(* IEC 61131-3 sources: Versio-VersionControlSystem/fixtures/projects/TC3_PlcSample_reStrText/TC3_PlcSample_reStrText/LibraryDocumentationSample Project/LibPOUs/B_DocuElements/Images, 1 file *)

(* ---- FB_Libdoc_Images.st ---- *)
(*

**Absolute or relative file path as directive argument**

Absolute path

.. image:: C:\Tc3LibDocImages\tulpis.jpg
   :width: 70px

Relative path

.. image:: ../../LibPics/penguins.jpg
   :width: 70px

**Left aligned image**

.. image:: ../../LibPics/desert.jpg
   :width: 20%

Description of the function block. Description of the function block. Description of the function block.
Description of the function block. Description of the function block. Description of the function block.
Description of the function block. Description of the function block. Description of the function block.
Description of the function block. Description of the function block. Description of the function block.

**Floating image, left aligned**

.. image:: ../../LibPics/desert.jpg
   :width: 20%
   :align: left

Description of the function block. Description of the function block. Description of the function block.
Description of the function block. Description of the function block. Description of the function block.
Description of the function block. Description of the function block. Description of the function block.
Description of the function block. Description of the function block. Description of the function block.

|
|
|
|
|

**Floating image, right aligned**

.. image:: ../../LibPics/desert.jpg
   :width: 20%
   :align: right

Description of the function block. Description of the function block. Description of the function block.
Description of the function block. Description of the function block. Description of the function block.
Description of the function block. Description of the function block. Description of the function block.
Description of the function block. Description of the function block. Description of the function block.

*)

FUNCTION_BLOCK FB_Libdoc_Images
VAR_INPUT
    nVarA : INT;
    nVarB : INT;
END_VAR
VAR_OUTPUT
    nSum : INT;
END_VAR
VAR
END_VAR
